Universal Robots URScript: T006_codellama_34b_baseline_rep2.urscript

def pick_and_place(bin_pose):
    # Home position
    movej(p[0, 0, 0, 0, 0, 0], v=350.0)

    # Above bin
    movel(p[0, 0, 120, 0, 0, 0], v=350.0)

    # Descend
